// TIA Portal V16 export
// export: Created 2000-01-01T00:00:00.0000000Z, ExportSetting None
FUNCTION "FC_Rung" : Void   // FC42, LAD
{ S7_Optimized_Access := 'TRUE' }
   VAR_INPUT
      Local : Int;
   END_VAR
BEGIN

REGION Network 1
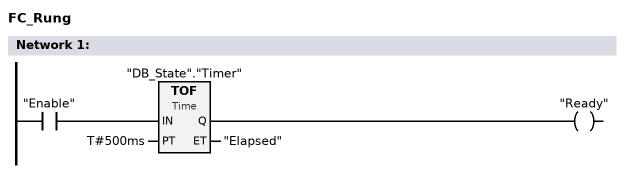
   RUNG wire#powerrail
      Contact( "Enable" )
      { S7_Templates := "time_type := Time" } "DB_State"."Timer".TOF(pt := T#500ms, et => "Elapsed")
      Coil( "Ready" )
   END_RUNG
   // the same network as SCL:
   "DB_State"."Timer".TOF(IN := "Enable", PT := T#500ms, ET => "Elapsed");
   "Ready" := "DB_State"."Timer".Q;
END_REGION
END_FUNCTION
